(* PLC project Conveyor_Sorting_System, CODESYS GmbH CODESYS CODESYS V3.5 SP20 *)
(* stored: creationDateTime 2026-10-27T11:30:00, modificationDateTime 2026-10-27T11:30:00 *)

TYPE E_OperationMode : (MODE_NONE := 0, MODE_MANUAL := 1, MODE_AUTOMATIC := 2);
END_TYPE

TYPE E_ObjectType : (OBJ_NONE := 0, OBJ_METAL := 1, OBJ_PLASTIC := 2, OBJ_DEFECTIVE := 3);
END_TYPE

TYPE E_SystemState : (STATE_IDLE := 0, STATE_RUNNING := 1, STATE_STOPPING := 2, STATE_ESTOP := 3, STATE_FAULT := 4);
END_TYPE

TYPE ST_BinStatus : STRUCT
  nCount : INT;
  nMaxCapacity : INT;
  bFull : BOOL;
END_STRUCT;
END_TYPE

PROGRAM PRG_Conveyor
  VAR
    tonDetectionFilter : TON;
    tDebounceTime : TIME := T#150MS;
    tonDelayToBin1 : TON;
    tTravelTimeBin1 : TIME := T#1650MS;
    tonDelayToBin2 : TON;
    tTravelTimeBin2 : TIME := T#3300MS;
    tpPusher1Actuate : TP;
    tPusher1PulseWidth : TIME := T#1200MS;
    tpPusher2Actuate : TP;
    tPusher2PulseWidth : TIME := T#1200MS;
    tpEntryAlert : TP;
    tEntryPulseWidth : TIME := T#500MS;
    tofMotorControlledStop : TOF;
    tRunoutDuration : TIME := T#3000MS;
    rtrigStart : R_TRIG;
    rtrigPusher1Fired : R_TRIG;
    rtrigPusher2Fired : R_TRIG;
    rtrigObjectAtBin3 : R_TRIG;
    rtrigSpawn : R_TRIG;
    bRawObjectDetected : BOOL := FALSE;
    bTargetBin1Armed : BOOL := FALSE;
    bTargetBin2Armed : BOOL := FALSE;
    bAutoPusher1Cmd : BOOL := FALSE;
    bAutoPusher2Cmd : BOOL := FALSE;
    tCurrentCycleTime : TIME;
    tLastCycleTime : TIME;
    rDeltaTime : REAL := 0.02;
    bCycleInitDone : BOOL := FALSE;
    rBeltLength : REAL := 1000.0;
    rSpawnIntervalTimer : REAL := 0.0;
    iSpawnSequenceCounter : INT := 1;
  END_VAR

            
// 1. CYCLE TIME CALCULATION
tCurrentCycleTime := TIME();
IF NOT bCycleInitDone THEN
    tLastCycleTime := tCurrentCycleTime;
    bCycleInitDone := TRUE;
    rDeltaTime := 0.02;
ELSE
    rDeltaTime := TIME_TO_REAL(tCurrentCycleTime - tLastCycleTime) / 1000.0;
    IF rDeltaTime <= 0.001 OR rDeltaTime > 0.1 THEN
        rDeltaTime := 0.02;
    END_IF;
    tLastCycleTime := tCurrentCycleTime;
END_IF;

// 2. OPERATING MODE DECODING & INTERLOCKING
IF GVL.iModeSelection = 1 THEN
    GVL.bModeManualActive := TRUE;
    GVL.bModeAutoActive   := FALSE;
ELSE
    GVL.iModeSelection    := 2;
    GVL.bModeManualActive := FALSE;
    GVL.bModeAutoActive   := TRUE;
END_IF;

// 3. LATCHING CIRCUIT FOR START / STOP
rtrigStart(CLK := GVL.bStartBtn);

IF GVL.bEmergencyStop THEN
    GVL.bRunLatch := FALSE;
    GVL.sSystemStatusMessage := 'EMERGENCY STOP ENGAGED! System halted.';
ELSIF GVL.bStopBtn THEN
    GVL.bRunLatch := FALSE;
    GVL.sSystemStatusMessage := 'Stop requested. Controlled deceleration in progress.';
ELSIF rtrigStart.Q THEN
    IF NOT GVL.bAlarmActive THEN
        GVL.bRunLatch := TRUE;
        GVL.sSystemStatusMessage := 'System Running - Conveyor Active.';
    ELSE
        GVL.sSystemStatusMessage := 'Cannot start: Clear active alarms first!';
    END_IF;
END_IF;

IF GVL.bResetFaultBtn THEN
    GVL.bAlarmActive            := FALSE;
    GVL.bInterlockBinFull       := FALSE;
    GVL.bInterlockPusherBlocked := FALSE;
    GVL.stBin1.bFull            := FALSE;
    GVL.stBin2.bFull            := FALSE;
    GVL.stBin3.bFull            := FALSE;
    GVL.stBin1.nCount           := 0;
    GVL.stBin2.nCount           := 0;
    GVL.stBin3.nCount           := 0;
    GVL.iTotalSorted            := 0;
    GVL.sSystemStatusMessage    := 'Alarms & Bin counts reset. System ready.';
END_IF;

// 4. CONTROLLED STOPPING USING TOF TIMER
tofMotorControlledStop(IN := GVL.bRunLatch, PT := tRunoutDuration);

IF GVL.bEmergencyStop THEN
    GVL.bMotorRun := FALSE;
    GVL.rConveyorSpeed := 0.0;
ELSIF GVL.bModeAutoActive THEN
    GVL.bMotorRun := tofMotorControlledStop.Q;
    IF GVL.bMotorRun THEN
        GVL.rConveyorSpeed := GVL.rSetSpeed;
    ELSE
        GVL.rConveyorSpeed := 0.0;
    END_IF;
ELSIF GVL.bModeManualActive THEN
    GVL.bMotorRun := GVL.bManualJogFwd;
    IF GVL.bMotorRun THEN
        GVL.rConveyorSpeed := GVL.rSetSpeed * 0.6;
    ELSE
        GVL.rConveyorSpeed := 0.0;
    END_IF;
END_IF;

// 5. OBJECT SPAWNING & CONVEYOR SIMULATION
rtrigSpawn(CLK := GVL.bSpawnNewObjectBtn);

IF GVL.bModeAutoActive AND GVL.bMotorRun AND NOT GVL.bObjectPresent THEN
    rSpawnIntervalTimer := rSpawnIntervalTimer + rDeltaTime;
    IF rSpawnIntervalTimer >= 1.5 THEN
        GVL.bObjectPresent := TRUE;
        GVL.rObjectPos := 0.0;
        GVL.iCurrentObjectType := iSpawnSequenceCounter;
        iSpawnSequenceCounter := iSpawnSequenceCounter + 1;
        IF iSpawnSequenceCounter > 3 THEN
            iSpawnSequenceCounter := 1;
        END_IF;
        rSpawnIntervalTimer := 0.0;
    END_IF;
ELSIF rtrigSpawn.Q AND NOT GVL.bObjectPresent THEN
    GVL.bObjectPresent := TRUE;
    GVL.rObjectPos := 0.0;
    GVL.iCurrentObjectType := GVL.iNextObjectTypeSelect;
    IF GVL.iCurrentObjectType < 1 OR GVL.iCurrentObjectType > 3 THEN
        GVL.iCurrentObjectType := 1;
    END_IF;
END_IF;

IF GVL.bObjectPresent AND GVL.bMotorRun THEN
    GVL.rObjectPos := GVL.rObjectPos + (GVL.rConveyorSpeed * rDeltaTime);
END_IF;

IF GVL.rObjectPos > rBeltLength THEN
    GVL.rObjectPos := rBeltLength;
END_IF;

// 6. SENSOR SIMULATION & DETECTION (TON Debounce)
GVL.bSensorEntry := GVL.bObjectPresent AND (GVL.rObjectPos >= 90.0 AND GVL.rObjectPos <= 140.0);

IF GVL.bObjectPresent AND (GVL.rObjectPos >= 230.0 AND GVL.rObjectPos <= 270.0) THEN
    bRawObjectDetected := TRUE;
    GVL.bSensorMetal   := (GVL.iCurrentObjectType = 1);
    GVL.bSensorHeight  := (GVL.iCurrentObjectType = 2);
ELSE
    bRawObjectDetected := FALSE;
    GVL.bSensorMetal   := FALSE;
    GVL.bSensorHeight  := FALSE;
END_IF;

GVL.bSensorBin1Station := GVL.bObjectPresent AND (GVL.rObjectPos >= 480.0 AND GVL.rObjectPos <= 520.0);
GVL.bSensorBin2Station := GVL.bObjectPresent AND (GVL.rObjectPos >= 730.0 AND GVL.rObjectPos <= 770.0);
GVL.bSensorBin3Station := GVL.bObjectPresent AND (GVL.rObjectPos >= 930.0 AND GVL.rObjectPos <= 970.0);

tonDetectionFilter(IN := bRawObjectDetected, PT := tDebounceTime);
GVL.bSensorDetectFiltered := tonDetectionFilter.Q;

IF GVL.bSensorDetectFiltered AND GVL.bModeAutoActive THEN
    IF GVL.iCurrentObjectType = 1 THEN
        bTargetBin1Armed := TRUE;
    ELSIF GVL.iCurrentObjectType = 2 THEN
        bTargetBin2Armed := TRUE;
    END_IF;
END_IF;

tpEntryAlert(IN := GVL.bSensorEntry, PT := tEntryPulseWidth);

// 7. SORTING DELAYS USING TON TIMERS
tonDelayToBin1(IN := bTargetBin1Armed AND GVL.bMotorRun, PT := tTravelTimeBin1);
tonDelayToBin2(IN := bTargetBin2Armed AND GVL.bMotorRun, PT := tTravelTimeBin2);

IF tonDelayToBin1.Q THEN
    bAutoPusher1Cmd  := TRUE;
    bTargetBin1Armed := FALSE;
END_IF;

IF tonDelayToBin2.Q THEN
    bAutoPusher2Cmd  := TRUE;
    bTargetBin2Armed := FALSE;
END_IF;

// 8. INTERLOCKING LOGIC
IF NOT GVL.bMotorRun THEN
    IF GVL.bManualPusher1 OR GVL.bManualPusher2 OR bAutoPusher1Cmd OR bAutoPusher2Cmd THEN
        GVL.bInterlockPusherBlocked := TRUE;
    END_IF;
    bAutoPusher1Cmd := FALSE;
    bAutoPusher2Cmd := FALSE;
ELSE
    GVL.bInterlockPusherBlocked := FALSE;
END_IF;

IF GVL.stBin1.nCount >= GVL.stBin1.nMaxCapacity THEN
    GVL.stBin1.bFull := TRUE;
    bAutoPusher1Cmd := FALSE;
    GVL.bInterlockBinFull := TRUE;
    GVL.bAlarmActive := TRUE;
    GVL.sSystemStatusMessage := 'ALARM: Bin 1 is FULL!';
END_IF;

IF GVL.stBin2.nCount >= GVL.stBin2.nMaxCapacity THEN
    GVL.stBin2.bFull := TRUE;
    bAutoPusher2Cmd := FALSE;
    GVL.bInterlockBinFull := TRUE;
    GVL.bAlarmActive := TRUE;
    GVL.sSystemStatusMessage := 'ALARM: Bin 2 is FULL!';
END_IF;

IF GVL.stBin3.nCount >= GVL.stBin3.nMaxCapacity THEN
    GVL.stBin3.bFull := TRUE;
    GVL.bInterlockBinFull := TRUE;
    GVL.bAlarmActive := TRUE;
    GVL.sSystemStatusMessage := 'ALARM: Reject Bin 3 is FULL!';
END_IF;

// 9. PUSHER ACTUATION USING TP TIMERS
tpPusher1Actuate(
    IN := (bAutoPusher1Cmd OR (GVL.bModeManualActive AND GVL.bManualPusher1)) 
          AND GVL.bMotorRun 
          AND NOT GVL.bPusher2 
          AND NOT GVL.stBin1.bFull 
          AND NOT GVL.bEmergencyStop,
    PT := tPusher1PulseWidth
);
GVL.bPusher1 := tpPusher1Actuate.Q;
IF GVL.bPusher1 THEN
    bAutoPusher1Cmd := FALSE;
END_IF;

tpPusher2Actuate(
    IN := (bAutoPusher2Cmd OR (GVL.bModeManualActive AND GVL.bManualPusher2)) 
          AND GVL.bMotorRun 
          AND NOT GVL.bPusher1 
          AND NOT GVL.stBin2.bFull 
          AND NOT GVL.bEmergencyStop,
    PT := tPusher2PulseWidth
);
GVL.bPusher2 := tpPusher2Actuate.Q;
IF GVL.bPusher2 THEN
    bAutoPusher2Cmd := FALSE;
END_IF;

// 10. PRODUCT SORTING EXECUTION & BIN ACCOUNTING
rtrigPusher1Fired(CLK := GVL.bPusher1);
rtrigPusher2Fired(CLK := GVL.bPusher2);
rtrigObjectAtBin3(CLK := (GVL.rObjectPos >= 950.0 AND GVL.bObjectPresent));

IF rtrigPusher1Fired.Q AND GVL.bObjectPresent AND (GVL.rObjectPos >= 450.0 AND GVL.rObjectPos <= 550.0) THEN
    GVL.stBin1.nCount  := GVL.stBin1.nCount + 1;
    GVL.iTotalSorted   := GVL.iTotalSorted + 1;
    GVL.bObjectPresent := FALSE;
    GVL.rObjectPos     := 0.0;
    bTargetBin1Armed   := FALSE;
    GVL.sSystemStatusMessage := 'Object (Metal) sorted into Bin 1 successfully.';
END_IF;

IF rtrigPusher2Fired.Q AND GVL.bObjectPresent AND (GVL.rObjectPos >= 700.0 AND GVL.rObjectPos <= 800.0) THEN
    GVL.stBin2.nCount  := GVL.stBin2.nCount + 1;
    GVL.iTotalSorted   := GVL.iTotalSorted + 1;
    GVL.bObjectPresent := FALSE;
    GVL.rObjectPos     := 0.0;
    bTargetBin2Armed   := FALSE;
    GVL.sSystemStatusMessage := 'Object (Plastic) sorted into Bin 2 successfully.';
END_IF;

IF rtrigObjectAtBin3.Q THEN
    GVL.stBin3.nCount  := GVL.stBin3.nCount + 1;
    GVL.iTotalSorted   := GVL.iTotalSorted + 1;
    GVL.bObjectPresent := FALSE;
    GVL.rObjectPos     := 0.0;
    bTargetBin1Armed   := FALSE;
    bTargetBin2Armed   := FALSE;
    IF GVL.iCurrentObjectType = 3 THEN
        GVL.sSystemStatusMessage := 'Defective item ejected to Bin 3 (Reject).';
    ELSE
        GVL.sSystemStatusMessage := 'Item passed through to Bin 3.';
    END_IF;
END_IF;

// 11. VISUALIZATION COORDINATES & COLOR BINDING
GVL.rVisuObjectX       := 120.0 + (GVL.rObjectPos * 0.6);
GVL.bVisuObjectVisible := GVL.bObjectPresent;

CASE GVL.iCurrentObjectType OF
    1: GVL.dwVisuObjectColor := 16#FF9E9E9E; // Metal (Gray)
    2: GVL.dwVisuObjectColor := 16#FF2196F3; // Plastic (Blue)
    3: GVL.dwVisuObjectColor := 16#FFE91E63; // Defective (Red)
ELSE
    GVL.dwVisuObjectColor := 16#FFFFFFFF;
END_CASE;

            
          
END_PROGRAM

CONFIGURATION Configuration
  VAR_GLOBAL  (* GVL *)
    bStartBtn : BOOL := FALSE;
    bStopBtn : BOOL := FALSE;
    bEmergencyStop : BOOL := FALSE;
    bResetFaultBtn : BOOL := FALSE;
    iModeSelection : INT := 2;
    bModeManualActive : BOOL;
    bModeAutoActive : BOOL;
    bManualJogFwd : BOOL := FALSE;
    bManualPusher1 : BOOL := FALSE;
    bManualPusher2 : BOOL := FALSE;
    bRunLatch : BOOL := FALSE;
    bMotorRun : BOOL := FALSE;
    rConveyorSpeed : REAL := 0.0;
    rSetSpeed : REAL := 150.0;
    rObjectPos : REAL := 0.0;
    iCurrentObjectType : INT := 1;
    bObjectPresent : BOOL := FALSE;
    iNextObjectTypeSelect : INT := 1;
    bSpawnNewObjectBtn : BOOL := FALSE;
    bSensorEntry : BOOL := FALSE;
    bSensorDetectFiltered : BOOL := FALSE;
    bSensorMetal : BOOL := FALSE;
    bSensorHeight : BOOL := FALSE;
    bSensorBin1Station : BOOL := FALSE;
    bSensorBin2Station : BOOL := FALSE;
    bSensorBin3Station : BOOL := FALSE;
    bPusher1 : BOOL := FALSE;
    bPusher2 : BOOL := FALSE;
    stBin1 : ST_BinStatus;
    stBin2 : ST_BinStatus;
    stBin3 : ST_BinStatus;
    iTotalSorted : INT := 0;
    bInterlockPusherBlocked : BOOL := FALSE;
    bInterlockBinFull : BOOL := FALSE;
    bAlarmActive : BOOL := FALSE;
    sSystemStatusMessage : STRING(80);
    rVisuObjectX : REAL := 120.0;
    rVisuObjectY : REAL := 220.0;
    bVisuObjectVisible : BOOL := FALSE;
    dwVisuObjectColor : DWORD := 16#FF9E9E9E;
  END_VAR
END_CONFIGURATION
